Fanuc KAREL source: KT00138.KL

PROGRAM KT00138
%NOLOCKGROUP
VAR
  R1: REAL
  I2: INTEGER
  OUT: REAL
BEGIN
  R1 = 2.0
    I2 = 3
  OUT = R1 DIV I2
END KT00138
